ABB RAPID module: WeldingAddin.mod

%%%
  VERSION:1
  LANGUAGE:ENGLISH
%%%
MODULE MOD_WeldingAddin

    ! -------------------------------
    ! Define customized variables here
    ! ...

	! Tool variables:
	PERS tooldata Tool1 := [TRUE,[[129.073,0.000,85.477],[0.98018657,0.00000000,0.19807649,0.00000000]],[1,[0,0,20],[1,0,0,0],0,0,0.005]];

	! Reference variables:
	PERS wobjdata RobotBase := [FALSE, TRUE, "", [[0,0,0],[1,0,0,0]],[[0.000,0.000,0.000],[1.00000000,0.00000000,0.00000000,0.00000000]]];

	PROC Main()
		ConfJ \On;
		ConfL \Off;
		! Program generated by RoboDK v5.7.3 for RoboDK Industrial on 02/07/2024 19:37:37
		! Using nominal kinematics.
		ArcLEnd None,v500,seam_end,weld_end,\Weave:=wv_end,z1,tool0 \WObj:=wobj0;
		MoveAbsJ [[-0.000001,0.000000,0.000000,0.000000,0.000000,-0.000000],[9E+09,9E+09,9E+09,9E+09,9E+09,9E+09]],v500,z1,Tool1 \WObj:=RobotBase;
		MoveAbsJ [[0.000000,3.211240,-15.423700,0.000000,12.212500,-0.000000],[9E+09,9E+09,9E+09,9E+09,9E+09,9E+09]],v500,z1,Tool1 \WObj:=RobotBase;
		ArcLStart [[1015.000,0.000,1272.000],[0.70710678,0.00000000,0.70710678,0.00000001],[0,0,0,1],[9E+09,9E+09,9E+09,9E+09,9E+09,9E+09]],v500,seam_start,weld_start,\Weave:=wv_start,z1,Tool1 \WObj:=RobotBase;
		ArcLEnd [[1015.000,0.000,1272.000],[0.70710678,0.00000000,0.70710678,0.00000001],[0,0,0,1],[9E+09,9E+09,9E+09,9E+09,9E+09,9E+09]],v500,seam_end,weld_end,\Weave:=wv_end,z1,Tool1 \WObj:=RobotBase;
		MoveAbsJ [[-0.000001,0.000000,0.000000,0.000000,0.000000,-0.000000],[9E+09,9E+09,9E+09,9E+09,9E+09,9E+09]],v500,z1,Tool1 \WObj:=RobotBase;
		! Previous line is a comment!
		ArcLEnd None,v500,seam_end,weld_end,\Weave:=wv_end,z1,Tool1 \WObj:=RobotBase;
		MoveAbsJ [[-0.000001,0.000000,0.000000,0.000000,0.000000,-0.000000],[9E+09,9E+09,9E+09,9E+09,9E+09,9E+09]],v500,z1,Tool1 \WObj:=RobotBase;
		! Previous line is a comment!
		MoveAbsJ [[0.000000,3.211240,-15.423700,0.000000,12.212500,-0.000000],[9E+09,9E+09,9E+09,9E+09,9E+09,9E+09]],v500,z1,Tool1 \WObj:=RobotBase;
		ArcLStart [[1015.000,0.000,1272.000],[0.70710678,0.00000000,0.70710678,0.00000001],[0,0,0,1],[9E+09,9E+09,9E+09,9E+09,9E+09,9E+09]],v500,seam_start,weld_start,\Weave:=wv_start,z1,Tool1 \WObj:=RobotBase;
		! Previous line is a comment!
		ArcLEnd [[1015.000,0.000,1272.000],[0.70710678,0.00000000,0.70710678,0.00000001],[0,0,0,1],[9E+09,9E+09,9E+09,9E+09,9E+09,9E+09]],v500,seam_end,weld_end,\Weave:=wv_end,z1,Tool1 \WObj:=RobotBase;
		! Previous line is a comment!
		MoveAbsJ [[-0.000001,0.000000,0.000000,0.000000,0.000000,-0.000000],[9E+09,9E+09,9E+09,9E+09,9E+09,9E+09]],v500,z1,Tool1 \WObj:=RobotBase;
	ENDPROC

ENDMODULE
